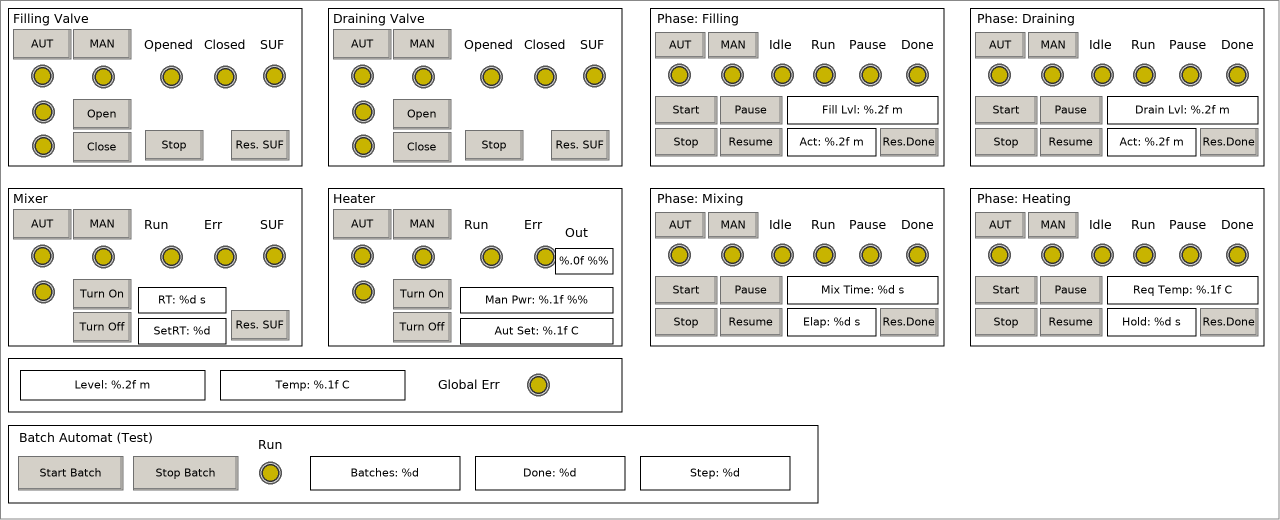
VISUALIZATION Visualization  // 1280x520
    Rectangle (8,8 294x158)
    Button (13,29 58x30), "AUT"
        OnMouseClick: toggle Global.Tank1.ValveFilling.Cmd.AutCtrl
    Button (73,29 58x30), "MAN"
        OnMouseClick: toggle Global.Tank1.ValveFilling.Cmd.ManCtrl
    Label (10,10 96x18), "Filling Valve"
    Button (73,99 58x30), "Open"
        OnMouseClick: toggle Global.Tank1.ValveFilling.Cmd.OpenMan
    Button (73,132 58x30), "Close"
        OnMouseClick: toggle Global.Tank1.ValveFilling.Cmd.CloseMan
    Lamp1 (29,63 27x26), variable: Global.Tank1.ValveFilling.State.AutCtrl, style: Lamp-Lamp1-Yellow
    Lamp1 (90,64 27x26), variable: Global.Tank1.ValveFilling.State.ManCtrl, style: Lamp-Lamp1-Yellow
    Lamp1 (158,64 27x26), variable: Global.Tank1.ValveFilling.State.Open, style: Lamp-Lamp1-Yellow
    Lamp1 (212,64 27x26), variable: Global.Tank1.ValveFilling.State.Closed, style: Lamp-Lamp1-Yellow
    Lamp1 (261,63 27x26), variable: Global.Tank1.ValveFilling.State.StartupFail, style: Lamp-Lamp1-Yellow
    Button (231,130 58x30), "Res. SUF"
        OnMouseClick: toggle Global.Tank1.ValveFilling.Cmd.ResetSUF
    Label (141,36 53x18), "Opened"
    Label (201,36 53x18), "Closed"
    Label (257,36 33x18), "SUF"
    Lamp1 (30,99 27x26), variable: Global.Tank1.ValveFilling.State.OpenOut, style: Lamp-Lamp1-Yellow
    Lamp1 (30,133 27x26), variable: Global.Tank1.ValveFilling.State.CloseOut, style: Lamp-Lamp1-Yellow
    Button (145,130 58x30), "Stop"
        OnMouseClick: toggle Global.Tank1.ValveFilling.Cmd.StopMan
    Rectangle (328,8 294x158)
    Button (333,29 58x30), "AUT"
        OnMouseClick: toggle Global.Tank1.ValveDraining.Cmd.AutCtrl
    Button (393,29 58x30), "MAN"
        OnMouseClick: toggle Global.Tank1.ValveDraining.Cmd.ManCtrl
    Label (330,10 120x18), "Draining Valve"
    Button (393,99 58x30), "Open"
        OnMouseClick: toggle Global.Tank1.ValveDraining.Cmd.OpenMan
    Button (393,132 58x30), "Close"
        OnMouseClick: toggle Global.Tank1.ValveDraining.Cmd.CloseMan
    Lamp1 (349,63 27x26), variable: Global.Tank1.ValveDraining.State.AutCtrl, style: Lamp-Lamp1-Yellow
    Lamp1 (410,64 27x26), variable: Global.Tank1.ValveDraining.State.ManCtrl, style: Lamp-Lamp1-Yellow
    Lamp1 (478,64 27x26), variable: Global.Tank1.ValveDraining.State.Open, style: Lamp-Lamp1-Yellow
    Lamp1 (532,64 27x26), variable: Global.Tank1.ValveDraining.State.Closed, style: Lamp-Lamp1-Yellow
    Lamp1 (581,63 27x26), variable: Global.Tank1.ValveDraining.State.StartupFail, style: Lamp-Lamp1-Yellow
    Button (551,130 58x30), "Res. SUF"
        OnMouseClick: toggle Global.Tank1.ValveDraining.Cmd.ResetSUF
    Label (461,36 53x18), "Opened"
    Label (521,36 53x18), "Closed"
    Label (577,36 33x18), "SUF"
    Lamp1 (350,99 27x26), variable: Global.Tank1.ValveDraining.State.OpenOut, style: Lamp-Lamp1-Yellow
    Lamp1 (350,133 27x26), variable: Global.Tank1.ValveDraining.State.CloseOut, style: Lamp-Lamp1-Yellow
    Button (465,130 58x30), "Stop"
        OnMouseClick: toggle Global.Tank1.ValveDraining.Cmd.StopMan
    Rectangle (8,188 294x158)
    Button (13,209 58x30), "AUT"
        OnMouseClick: toggle Global.Tank1.Mixer.Cmd.AutCtrl
    Button (73,209 58x30), "MAN"
        OnMouseClick: toggle Global.Tank1.Mixer.Cmd.ManCtrl
    Label (10,190 96x18), "Mixer"
    Button (73,279 58x30), "Turn On"
        OnMouseClick: toggle Global.Tank1.Mixer.Cmd.TurnOnMan
    Button (73,312 58x30), "Turn Off"
        OnMouseClick: toggle Global.Tank1.Mixer.Cmd.TurnOffMan
    Lamp1 (29,243 27x26), variable: Global.Tank1.Mixer.State.AutCtrl, style: Lamp-Lamp1-Yellow
    Lamp1 (90,244 27x26), variable: Global.Tank1.Mixer.State.ManCtrl, style: Lamp-Lamp1-Yellow
    Lamp1 (158,244 27x26), variable: Global.Tank1.Mixer.State.Run, style: Lamp-Lamp1-Yellow
    Lamp1 (212,244 27x26), variable: Global.Tank1.Mixer.State.GenErr, style: Lamp-Lamp1-Yellow
    Lamp1 (261,243 27x26), variable: Global.Tank1.Mixer.State.StartUpFail, style: Lamp-Lamp1-Yellow
    Button (231,310 58x30), "Res. SUF"
        OnMouseClick: toggle Global.Tank1.Mixer.Cmd.ResetSUF
    Label (141,216 53x18), "Run"
    Label (201,216 53x18), "Err"
    Label (257,216 33x18), "SUF"
    Lamp1 (30,279 27x26), variable: Global.Tank1.Mixer.State.RunOut, style: Lamp-Lamp1-Yellow
    Rectangle (328,188 294x158)
    Button (333,209 58x30), "AUT"
        OnMouseClick: toggle Global.Tank1.Heater.Cmd.AutCtrl
    Button (393,209 58x30), "MAN"
        OnMouseClick: toggle Global.Tank1.Heater.Cmd.ManCtrl
    Label (330,190 96x18), "Heater"
    Button (393,279 58x30), "Turn On"
        OnMouseClick: toggle Global.Tank1.Heater.Cmd.TurnOnMan
    Button (393,312 58x30), "Turn Off"
        OnMouseClick: toggle Global.Tank1.Heater.Cmd.TurnOffMan
    Lamp1 (349,243 27x26), variable: Global.Tank1.Heater.State.AutCtrl, style: Lamp-Lamp1-Yellow
    Lamp1 (410,244 27x26), variable: Global.Tank1.Heater.State.ManCtrl, style: Lamp-Lamp1-Yellow
    Lamp1 (478,244 27x26), variable: Global.Tank1.Heater.State.EnableOut, style: Lamp-Lamp1-Yellow
    Lamp1 (532,244 27x26), variable: Global.Tank1.Heater.State.GenErr, style: Lamp-Lamp1-Yellow
    Label (461,216 53x18), "Run"
    Label (521,216 53x18), "Err"
    Lamp1 (350,279 27x26), variable: Global.Tank1.Heater.State.EnableOut, style: Lamp-Lamp1-Yellow
    Rectangle (138,287 88x26), "RT: %d s", text variable: Global.Tank1.Mixer.State.RT
    Rectangle (138,318 88x26), "SetRT: %d", text variable: Global.Tank1.Mixer.Cmd.SetRT
        OnMouseClick: write the text variable via Default
    Label (562,224 45x18), "Out"
    Rectangle (555,248 58x26), "%.0f %%", text variable: Global.Tank1.Heater.State.HeatingOut
    Rectangle (460,287 153x26), "Man Pwr: %.1f %%", text variable: Global.Tank1.Heater.ParamHeatingPowerManual
        OnMouseClick: write the text variable via Default
    Rectangle (460,318 153x26), "Aut Set: %.1f C", text variable: Global.Tank1.Heater.ParamHeatingSetPointAutomat
        OnMouseClick: write the text variable via Default
    Rectangle (8,358 614x54)
    Rectangle (20,370 185x30), "Level: %.2f m", text variable: Global.Tank1.Filling.WaterLevel
    Rectangle (220,370 185x30), "Temp: %.1f C", text variable: Global.Tank1.Heating.WaterTemp
    Label (435,376 85x20), "Global Err"
    Lamp1 (525,372 27x26), variable: Global.Tank1.GlobalError, style: Lamp-Lamp1-Yellow
    Rectangle (650,8 294x158)
    Label (654,10 140x18), "Phase: Filling"
    Button (655,32 50x26), "AUT"
        OnMouseClick: toggle Global.Tank1.Filling.Cmd.AutCtrl
    Button (708,32 50x26), "MAN"
        OnMouseClick: toggle Global.Tank1.Filling.Cmd.ManCtrl
    Label (766,36 38x18), "Idle"
    Label (808,36 38x18), "Run"
    Label (846,36 52x18), "Pause"
    Label (898,36 44x18), "Done"
    Lamp1 (666,62 27x26), variable: Global.Tank1.Filling.State.AutCtrl, style: Lamp-Lamp1-Yellow
    Lamp1 (719,62 27x26), variable: Global.Tank1.Filling.State.ManCtrl, style: Lamp-Lamp1-Yellow
    Lamp1 (769,62 27x26), variable: Global.Tank1.Filling.State.Idle, style: Lamp-Lamp1-Yellow
    Lamp1 (811,62 27x26), variable: Global.Tank1.Filling.State.Running, style: Lamp-Lamp1-Yellow
    Lamp1 (857,62 27x26), variable: Global.Tank1.Filling.State.Paused, style: Lamp-Lamp1-Yellow
    Lamp1 (904,62 27x26), variable: Global.Tank1.Filling.State.Done, style: Lamp-Lamp1-Yellow
    Button (655,96 62x28), "Start"
        OnMouseClick: toggle Global.Tank1.Filling.Cmd.StartMan
    Button (720,96 62x28), "Pause"
        OnMouseClick: toggle Global.Tank1.Filling.Cmd.PauseMan
    Button (655,128 62x28), "Stop"
        OnMouseClick: toggle Global.Tank1.Filling.Cmd.StopMan
    Button (720,128 62x28), "Resume"
        OnMouseClick: toggle Global.Tank1.Filling.Cmd.ResumeMan
    Rectangle (787,96 151x28), "Fill Lvl: %.2f m", text variable: Global.Tank1.Filling.ParamFillLevel
        OnMouseClick: write the text variable via Default
    Rectangle (787,128 89x28), "Act: %.2f m", text variable: Global.Tank1.Filling.WaterLevel
    Button (880,128 58x28), "Res.Done"
        OnMouseClick: toggle Global.Tank1.Filling.Cmd.ResetDone
    Rectangle (970,8 294x158)
    Label (974,10 140x18), "Phase: Draining"
    Button (975,32 50x26), "AUT"
        OnMouseClick: toggle Global.Tank1.Draining.Cmd.AutCtrl
    Button (1028,32 50x26), "MAN"
        OnMouseClick: toggle Global.Tank1.Draining.Cmd.ManCtrl
    Label (1086,36 38x18), "Idle"
    Label (1128,36 38x18), "Run"
    Label (1166,36 52x18), "Pause"
    Label (1218,36 44x18), "Done"
    Lamp1 (986,62 27x26), variable: Global.Tank1.Draining.State.AutCtrl, style: Lamp-Lamp1-Yellow
    Lamp1 (1039,62 27x26), variable: Global.Tank1.Draining.State.ManCtrl, style: Lamp-Lamp1-Yellow
    Lamp1 (1089,62 27x26), variable: Global.Tank1.Draining.State.Idle, style: Lamp-Lamp1-Yellow
    Lamp1 (1131,62 27x26), variable: Global.Tank1.Draining.State.Running, style: Lamp-Lamp1-Yellow
    Lamp1 (1177,62 27x26), variable: Global.Tank1.Draining.State.Paused, style: Lamp-Lamp1-Yellow
    Lamp1 (1224,62 27x26), variable: Global.Tank1.Draining.State.Done, style: Lamp-Lamp1-Yellow
    Button (975,96 62x28), "Start"
        OnMouseClick: toggle Global.Tank1.Draining.Cmd.StartMan
    Button (1040,96 62x28), "Pause"
        OnMouseClick: toggle Global.Tank1.Draining.Cmd.PauseMan
    Button (975,128 62x28), "Stop"
        OnMouseClick: toggle Global.Tank1.Draining.Cmd.StopMan
    Button (1040,128 62x28), "Resume"
        OnMouseClick: toggle Global.Tank1.Draining.Cmd.ResumeMan
    Rectangle (1107,96 151x28), "Drain Lvl: %.2f m", text variable: Global.Tank1.Draining.ParamDrainLevel
        OnMouseClick: write the text variable via Default
    Rectangle (1107,128 89x28), "Act: %.2f m", text variable: Global.Tank1.Draining.WaterLevel
    Button (1200,128 58x28), "Res.Done"
        OnMouseClick: toggle Global.Tank1.Draining.Cmd.ResetDone
    Rectangle (650,188 294x158)
    Label (654,190 140x18), "Phase: Mixing"
    Button (655,212 50x26), "AUT"
        OnMouseClick: toggle Global.Tank1.Mixing.Cmd.AutCtrl
    Button (708,212 50x26), "MAN"
        OnMouseClick: toggle Global.Tank1.Mixing.Cmd.ManCtrl
    Label (766,216 38x18), "Idle"
    Label (808,216 38x18), "Run"
    Label (846,216 52x18), "Pause"
    Label (898,216 44x18), "Done"
    Lamp1 (666,242 27x26), variable: Global.Tank1.Mixing.State.AutCtrl, style: Lamp-Lamp1-Yellow
    Lamp1 (719,242 27x26), variable: Global.Tank1.Mixing.State.ManCtrl, style: Lamp-Lamp1-Yellow
    Lamp1 (769,242 27x26), variable: Global.Tank1.Mixing.State.Idle, style: Lamp-Lamp1-Yellow
    Lamp1 (811,242 27x26), variable: Global.Tank1.Mixing.State.Running, style: Lamp-Lamp1-Yellow
    Lamp1 (857,242 27x26), variable: Global.Tank1.Mixing.State.Paused, style: Lamp-Lamp1-Yellow
    Lamp1 (904,242 27x26), variable: Global.Tank1.Mixing.State.Done, style: Lamp-Lamp1-Yellow
    Button (655,276 62x28), "Start"
        OnMouseClick: toggle Global.Tank1.Mixing.Cmd.StartMan
    Button (720,276 62x28), "Pause"
        OnMouseClick: toggle Global.Tank1.Mixing.Cmd.PauseMan
    Button (655,308 62x28), "Stop"
        OnMouseClick: toggle Global.Tank1.Mixing.Cmd.StopMan
    Button (720,308 62x28), "Resume"
        OnMouseClick: toggle Global.Tank1.Mixing.Cmd.ResumeMan
    Rectangle (787,276 151x28), "Mix Time: %d s", text variable: Global.Tank1.Mixing.ParamTimeSec
        OnMouseClick: write the text variable via Default
    Rectangle (787,308 89x28), "Elap: %d s", text variable: Global.Tank1.Mixing.ElapsedTimeSec
    Button (880,308 58x28), "Res.Done"
        OnMouseClick: toggle Global.Tank1.Mixing.Cmd.ResetDone
    Rectangle (970,188 294x158)
    Label (974,190 140x18), "Phase: Heating"
    Button (975,212 50x26), "AUT"
        OnMouseClick: toggle Global.Tank1.Heating.Cmd.AutCtrl
    Button (1028,212 50x26), "MAN"
        OnMouseClick: toggle Global.Tank1.Heating.Cmd.ManCtrl
    Label (1086,216 38x18), "Idle"
    Label (1128,216 38x18), "Run"
    Label (1166,216 52x18), "Pause"
    Label (1218,216 44x18), "Done"
    Lamp1 (986,242 27x26), variable: Global.Tank1.Heating.State.AutCtrl, style: Lamp-Lamp1-Yellow
    Lamp1 (1039,242 27x26), variable: Global.Tank1.Heating.State.ManCtrl, style: Lamp-Lamp1-Yellow
    Lamp1 (1089,242 27x26), variable: Global.Tank1.Heating.State.Idle, style: Lamp-Lamp1-Yellow
    Lamp1 (1131,242 27x26), variable: Global.Tank1.Heating.State.Running, style: Lamp-Lamp1-Yellow
    Lamp1 (1177,242 27x26), variable: Global.Tank1.Heating.State.Paused, style: Lamp-Lamp1-Yellow
    Lamp1 (1224,242 27x26), variable: Global.Tank1.Heating.State.Done, style: Lamp-Lamp1-Yellow
    Button (975,276 62x28), "Start"
        OnMouseClick: toggle Global.Tank1.Heating.Cmd.StartMan
    Button (1040,276 62x28), "Pause"
        OnMouseClick: toggle Global.Tank1.Heating.Cmd.PauseMan
    Button (975,308 62x28), "Stop"
        OnMouseClick: toggle Global.Tank1.Heating.Cmd.StopMan
    Button (1040,308 62x28), "Resume"
        OnMouseClick: toggle Global.Tank1.Heating.Cmd.ResumeMan
    Rectangle (1107,276 151x28), "Req Temp: %.1f C", text variable: Global.Tank1.Heating.ParamReqTemp
        OnMouseClick: write the text variable via Default
    Rectangle (1107,308 89x28), "Hold: %d s", text variable: Global.Tank1.Heating.fTime
    Button (1200,308 58x28), "Res.Done"
        OnMouseClick: toggle Global.Tank1.Heating.Cmd.ResetDone
    Rectangle (8,425 810x78)
    Label (16,429 180x20), "Batch Automat (Test)"
    Button (18,456 105x34), "Start Batch"
        OnMouseClick: toggle Test.bStartBatch
    Button (133,456 105x34), "Stop Batch"
        OnMouseClick: toggle Test.bStopBatch
    Label (255,436 38x18), "Run"
    Lamp1 (257,460 27x26), variable: Test.bRunning, style: Lamp-Lamp1-Yellow
    Rectangle (310,456 150x34), "Batches: %d", text variable: Test.nTargetBatches
        OnMouseClick: write the text variable via Default
    Rectangle (475,456 150x34), "Done: %d", text variable: Test.nCompletedBatches
    Rectangle (640,456 150x34), "Step: %d", text variable: Test.State
END_VISUALIZATION

(* stored: Version 1.1.0.1, ProductVersion 3.1.4026.21
   Visu Visualization: Id {a6343251-0068-49ba-9adb-31cb88a6e465} *)
